(* IEC 61131-3 sources: PLC-conveyor-testbench/plc/ConveyorController/pous/function-blocks, 3 files *)

(* ---- FB_Conveyor.st ---- *)
FUNCTION_BLOCK FB_Conveyor
VAR_INPUT
    xStart          : BOOL;
    xStop           : BOOL;
    xReset          : BOOL;
    xEmergencyStop  : BOOL;
    xJamDetected    : BOOL;
END_VAR

VAR_OUTPUT
    xMotorEnable    : BOOL := FALSE;
    iState          : INT := 0;
    iFaultCode      : INT := 0;
END_VAR

VAR
    fbStartEdge     : R_TRIG;
    fbResetEdge     : R_TRIG;
END_VAR

(* Detect operator command edges *)
fbStartEdge(CLK := xStart);
fbResetEdge(CLK := xReset);

(* Simulated emergency stop has highest priority *)
IF xEmergencyStop THEN

    iState := 2;
    iFaultCode := 2;

(* Handle latched fault *)
ELSIF iState = 2 THEN

    IF fbResetEdge.Q AND NOT xJamDetected THEN

        iState := 0;
        iFaultCode := 0;

    END_IF;

(* Handle conveyor jam *)
ELSIF xJamDetected AND (iState = 1) THEN

    iState := 2;
    iFaultCode := 1;

(* Normal operating states *)
ELSE

    CASE iState OF

        0:  (* IDLE *)

            IF fbStartEdge.Q AND NOT xStop THEN
                iState := 1;
            END_IF;

        1:  (* RUNNING *)

            IF xStop THEN
                iState := 0;
            END_IF;

        ELSE

            (* Invalid state *)
            iState := 2;
            iFaultCode := 3;

    END_CASE;

END_IF;

(* Motor command *)
xMotorEnable :=
    (iState = 1)
    AND NOT xStop
    AND NOT xEmergencyStop
    AND NOT xJamDetected;

END_FUNCTION_BLOCK

(* ---- FB_ItemTracker.st ---- *)
FUNCTION_BLOCK FB_ItemTracker
VAR_INPUT
    xRunEnable       : BOOL;
    xEntrySensor     : BOOL;
    xExitSensor      : BOOL;
END_VAR

VAR_OUTPUT
    xItemInTransit    : BOOL := FALSE;
    udiItemCount      : UDINT := 0;
END_VAR

VAR
    fbEntryEdge       : R_TRIG;
    fbExitEdge        : R_TRIG;
END_VAR

(* Detect sensor rising edges *)
fbEntryEdge(CLK := xEntrySensor);
fbExitEdge(CLK := xExitSensor);

(* Product tracking *)
IF xRunEnable THEN

    (* Complete an active transfer *)
    IF fbExitEdge.Q AND xItemInTransit THEN

        udiItemCount := udiItemCount + 1;
        xItemInTransit := FALSE;

    (* Register a new product *)
    ELSIF fbEntryEdge.Q AND NOT xItemInTransit THEN

        xItemInTransit := TRUE;

    END_IF;

ELSE

    (* Discard incomplete transfer when disabled *)
    xItemInTransit := FALSE;

END_IF;

END_FUNCTION_BLOCK

(* ---- FB_JamMonitor.st ---- *)
FUNCTION_BLOCK FB_JamMonitor
VAR_INPUT
    xEnable         : BOOL;
    xItemInTransit  : BOOL;
    tTimeout        : TIME := T#3s;
END_VAR

VAR_OUTPUT
    xJamDetected    : BOOL;
    tElapsed        : TIME;
END_VAR

VAR
    fbTimer         : TON;
END_VAR

(* Conveyor transfer timeout supervision *)

fbTimer(
    IN := xEnable AND xItemInTransit,
    PT := tTimeout
);

(* Output signals *)
xJamDetected := fbTimer.Q;
tElapsed := fbTimer.ET;

END_FUNCTION_BLOCK
